Fanuc KAREL source: KD00006.KL

PROGRAM KD00006
%NOLOCKGROUP
%NOPAUSESHFT
VAR
  I: INTEGER
  J: INTEGER
  B: BOOLEAN
  R: REAL
  S: STRING[80]
BEGIN
  I = 1
END KD00006
